Fanuc KAREL source: kt00908.KL

-- PROVISIONAL review KL for V1013-1; original PC SHA256 2d0b6ddd6f267498e48336c45e2d3749fe9ba6db8d1acbe6ea6de497c4fc2661
-- Incomplete behavior may be omitted. Consult companion uncertainty JSON. Do not deploy.
PROGRAM KT00908
%NOLOCKGROUP
BEGIN
  -- UNRESOLVED_PC offsets 5-28; opcodes 27,22,1C,31,4A
  -- UNRESOLVED_PC offsets 33-37; opcodes 7F
END KT00908
